// TIA Portal V20 export
// export: Created 2026-10-12T05:42:29.1445004Z, ExportSetting WithDefaults, DisplayName Totally Integrated Automation Portal, DisplayVersion V20, DisplayName TIA Portal Openness, DisplayVersion V20, DisplayName TIA Portal Teamcenter Gateway, DisplayVersion V20, DisplayName TIA Portal Version Control Interface, DisplayVersion V20, DisplayName SINAMICS Startdrive Advanced, DisplayVersion V20 SP1 Update 2, DisplayName SINAMICS Startdrive G110M, G120, G120C, G120D, G120P, G115D, DisplayVersion V20 SP1 Update 2, DisplayName SINAMICS Startdrive G130, G150, S120, S150, SINAMICS MV, G220, S200, S210, DisplayVersion V20 SP1 Update 2, DisplayName STEP 7 Professional, DisplayVersion V20, DisplayName STEP 7 Safety, DisplayVersion V20, DisplayName WinCC Basic/Comfort/Advanced, DisplayVersion V20, DisplayName WinCC Professional, DisplayVersion V20, DisplayName WinCC Unified, DisplayVersion V20
FUNCTION "FRK_AlarmBegin" : Void   // FC30, SCL
{ S7_Optimized_Access := 'TRUE' }
VERSION : 0.1
// stored: AutoNumber true, IsIECCheckEnabled false, SetENOAutomatically false, UDAEnableTagReadback false
   VAR_INPUT
      Startup : Bool;
   END_VAR
   VAR_IN_OUT
      AlarmLog : "FRK_AlarmLog";
   END_VAR
   VAR_TEMP
      Index : Int;
   END_VAR
BEGIN

   FOR #Index := 1 TO 16 DO
       #AlarmLog.Touched[#Index] := FALSE;
       IF #Startup THEN
           #AlarmLog.Active[#Index] := "FRK_UnitScratch".EmptyEvent;
           #AlarmLog.Automatic[#Index] := FALSE;
           #AlarmLog.ComeMs[#Index] := 0;
       END_IF;
   END_FOR;
   IF #Startup THEN
       FOR #Index := 1 TO 64 DO
           #AlarmLog.Ring[#Index] := "FRK_UnitScratch".EmptyEvent;
       END_FOR;
       #AlarmLog.RingHead := 0;
       #AlarmLog.RingUsed := 0;
       #AlarmLog.Truncated := FALSE;
   END_IF;
   "FRK_AlarmRefresh"(AlarmLog := #AlarmLog);
END_FUNCTION
